(* IEC 61131-3 sources: vscode-structured-text/test/format/fixtures, 10 files *)

(* ---- types.expected.st ---- *)
TYPE tComplex
(*
Copyright ©<Company>. All rights reserved.
*)
    STRUCT
        rRe : Real; //Complex real part
        rIm : Real; //Complex imaginary part
    END_STRUCT
END_TYPE

TYPE uMaCommand :
    UNION
        b : tMaCommand; //For Bit Access
        w : Word;       //For Word Access
    END_UNION
END_TYPE

TYPE eColor : (Red := 0, Green, Blue);
END_TYPE
TYPE tArr : Array[1..10] Of Pointer To Int;
END_TYPE

(* ---- types.input.st ---- *)
TYPE tComplex
(*
Copyright ©<Company>. All rights reserved.
*)
STRUCT
rRe : REAL ; //Complex real part
rIm : REAL ; //Complex imaginary part
END_STRUCT
END_TYPE

TYPE uMaCommand :
UNION
 b   : tMaCommand; //For Bit Access
 w   : WORD;  //For Word Access
END_UNION
END_TYPE

TYPE eColor : (Red := 0, Green, Blue); END_TYPE
TYPE tArr : ARRAY [1..10] OF POINTER TO INT; END_TYPE

(* ---- oneline.expected.st ---- *)
FUNCTION fcAdd : Int
VAR_INPUT
    a : Int;
    b : Int;
END_VAR
tiSourcIndex                            := tiSourcIndex + 1;
tiDestinationIndex                      := tiDestinationIndex + 1;
If xxx Then
    yyy                                 := 1;
End_If
fcAdd                                   := a + b;
END_FUNCTION

(* ---- oneline.input.st ---- *)
FUNCTION fcAdd : INT
VAR_INPUT a : INT; b : INT; END_VAR
tiSourcIndex := tiSourcIndex + 1; tiDestinationIndex := tiDestinationIndex + 1;
IF xxx THEN yyy := 1; END_IF
fcAdd:=a+b;
END_FUNCTION

(* ---- fbruntime.expected.st ---- *)
(*

**©2026 <Company> - TITLE =[V#01.01.01.03] Measures task runtime and jitter**

========================  ================  ===========  =========================================
Version Number            Date              Signature    Description
========================  ================  ===========  =========================================
V#01.01.01.03             2026.06.01        <Sign>         Original version.
========================  ================  ===========  =========================================
*)

FUNCTION_BLOCK fbRuntime
(*
Copyright ©2026 <Company>. All rights reserved.
AUTHOR : <Sign>
FAMILY : System
NAME   : fbRuntime
*)

VAR CONSTANT
    {attribute 'hide'} cliNsPerUs : LInt := 1000;      //Nanoseconds per microsecond
END_VAR

VAR_INPUT
    ibStart : Bool; //Start call
    ibReset : Bool; //Reset min and max
END_VAR

VAR_OUTPUT
    qltRuntime       : LTime; // Actual runtime
    qliRuntimeJitter : LInt;  // [us] Runtime jitter
    qltRuntimeMax    : LTime; // Maximum runtime
    qltRuntimemin    : LTime; // Minimum runtime
END_VAR

VAR //Static
    {attribute 'hide'} sltNow        : LTime;
    {attribute 'hide'} sltRuntimeMax : LTime;
END_VAR

VAR_TEMP
    {attribute 'hide'} tbRestart  : Bool;
    {attribute 'hide'} tltRuntime : LTime;
    {attribute 'hide'} tliJitter  : LInt;
    {attribute 'hide'} tltNow     : LTime;
END_VAR

//Populate Temporaries
tbRestart                               := gSystem.bRestart();
tltNow                                  := LTime();
tltRuntime                              := tltNow - sltNow;

//Handle restart and reset
If (ibReset Or tbRestart) Then
    sltRuntimeMax                       := LTime#0s;
    sltRuntimeMin                       := LTime#1d;
    sltNow                              := tltNow;
    Return;
End_If;

//Handle start and end call
If ibStart Then
    sltNow                              := tltNow;
    qltRuntime                          := Ltime#0s;
    qliRuntimeJitter                    := 0;
    Return;
End_If;

//Handle Min/Max cycle time
If (tltRuntime > sltRuntimeMax) Then
    sltRuntimeMax                       := tltRuntime;
Elsif (tltRuntime < sltRuntimeMin) Then
    sltRuntimeMin                       := tltRuntime;
End_If;
tliJitter                               := (LTime_To_LInt(tltRuntime) - sliJitter) / cliNsPerUs;
sliJitter                               := LTime_To_LInt(tltRuntime);

//Write to outputs
qltRuntime                              := tltRuntime;
qliRuntimeJitter                        := tliJitter; // jitter
qltRuntimeMax                           := sltRuntimeMax;
qltRuntimeMin                           := sltRuntimeMin;
END_FUNCTION_BLOCK

(* ---- fbruntime.input.st ---- *)
(*

**©2026 <Company> - TITLE =[V#01.01.01.03] Measures task runtime and jitter**

========================  ================  ===========  =========================================
Version Number            Date              Signature    Description
========================  ================  ===========  =========================================
V#01.01.01.03             2026.06.01        <Sign>         Original version.
========================  ================  ===========  =========================================
*)

FUNCTION_BLOCK fbRuntime
(*
Copyright ©2026 <Company>. All rights reserved.
AUTHOR : <Sign>
FAMILY : System
NAME   : fbRuntime
*)

VAR CONSTANT
{attribute 'hide'}     cliNsPerUs : Lint:= 1000;      //Nanoseconds per microsecond
END_VAR
VAR_INPUT
 ibStart    : Bool;        //Start call
 ibReset    : Bool;        //Reset min and max
END_VAR

VAR_OUTPUT
 qltRuntime   : LTime;  // Actual runtime
 qliRuntimeJitter  : Lint;         // [us] Runtime jitter
 qltRuntimeMax   : LTime;  // Maximum runtime
 qltRuntimemin   : LTime;  // Minimum runtime
END_VAR

VAR //Static
{attribute 'hide'}     sltNow  : LTime;
{attribute 'hide'}     sltRuntimeMax : LTime;
END_VAR

VAR_TEMP
{attribute 'hide'}     tbRestart : Bool;
{attribute 'hide'}     tltRuntime    : LTime;
{attribute 'hide'}     tliJitter    : Lint ;
{attribute 'hide'}     tltNow  : LTime;
END_VAR

//Populate Temporaries
tbRestart := gSystem.bRestart();
tltNow  := LTime();
tltRuntime := tltNow - sltNow;

//Handle restart and reset
IF (ibReset OR tbRestart) THEN
sltRuntimeMax := LTime#0s;
    sltRuntimeMin                  := LTime#1d;
      sltNow                        := tltNow;
    RETURN;
END_IF;

//Handle start and end call
If ibStart Then sltNow := tltNow; qltRuntime := Ltime#0s;
    qliRuntimeJitter            := 0;
    Return;
End_If;

//Handle Min/Max cycle time
If (tltRuntime > sltRuntimeMax) Then
    sltRuntimeMax                    := tltRuntime;
Elsif (tltRuntime < sltRuntimeMin) Then
    sltRuntimeMin                    := tltRuntime;
End_If;
tliJitter:=(LTIME_TO_LINT(tltRuntime)-sliJitter)/cliNsPerUs;
sliJitter                            := LTime_To_Lint(tltRuntime);

//Write to outputs
qltRuntime                          := tltRuntime;
qliRuntimeJitter            := tliJitter; // jitter
qltRuntimeMax              := sltRuntimeMax;
qltRuntimeMin               := sltRuntimeMin;
END_FUNCTION_BLOCK

(* ---- oop.expected.st ---- *)
{attribute 'qualified_only'}
INTERFACE iMotor EXTENDS iBase
METHOD mStart : Bool
VAR_INPUT
    ibForce : Bool;
END_VAR
END_METHOD
END_INTERFACE

FUNCTION_BLOCK PUBLIC fbMotor EXTENDS fbBase IMPLEMENTS iMotor
VAR_INPUT
    RX : Bool;   //Initialize filter
END_VAR;

VAR //Static Data
    sbRx   : Bool;   //Initialize filter
    sRef   : Reference To Int;
    spData : Pointer To tData;
END_VAR;

VAR_TEMP
    tbRx : Bool;    //Initialize filter
END_VAR;
BEGIN
tbRx                                    := RX And Not sbRx; //tbRx is positive edge for RX
sbRx                                    := RX;              //Save RX in sbRx to disable edge as long as RX stays true.
{IF defined (DEBUG)}
If tbRx Then
    This^.mLog(sMsg := 'edge');
End_If;
{END_IF}
spData                                  := __New(tData);
sRef REF= siValue;
If ((tbyXa And 16#01) <> 16#00) Then  //Test for positive edge on bit zero in the byte
    sbAlarm S= True;
End_If
METHOD PRIVATE mLog : Bool
VAR_INPUT
    sMsg : String(80);
END_VAR
mLog                                    := True;
END_METHOD

PROPERTY pbRunning : Bool
END_PROPERTY
END_FUNCTION_BLOCK

(* ---- oop.input.st ---- *)
{attribute 'qualified_only'}
INTERFACE iMotor EXTENDS iBase
METHOD mStart : BOOL
VAR_INPUT
ibForce : BOOL;
END_VAR
END_METHOD
END_INTERFACE

FUNCTION_BLOCK PUBLIC fbMotor EXTENDS fbBase IMPLEMENTS iMotor
VAR_INPUT
    RX   : Bool ;   //Initialize filter
END_VAR;
VAR //Static Data
    sbRx  : Bool ;   //Initialize filter
    sRef : REFERENCE TO INT;
    spData : POINTER TO tData;
END_VAR;
VAR_TEMP
    tbRx         : Bool ;    //Initialize filter
END_VAR;
BEGIN
tbRx   := RX And Not sbRx; //tbRx is positive edge for RX
sbRx   := RX;              //Save RX in sbRx to disable edge as long as RX stays true.
{IF defined (DEBUG)}
If tbRx Then
    THIS^.mLog(sMsg := 'edge');
End_If;
{END_IF}
spData := __NEW(tData);
sRef REF= siValue;
IF ((tbyXa AND 16#01) <> 16#00) THEN  //Test for positive edge on bit zero in the byte
    sbAlarm S= TRUE;
END_IF
METHOD PRIVATE mLog : BOOL
VAR_INPUT
    sMsg : STRING(80);
END_VAR
mLog := TRUE;
END_METHOD

PROPERTY pbRunning : BOOL
END_PROPERTY
END_FUNCTION_BLOCK

(* ---- fsm.expected.st ---- *)
VAR CONSTANT
    //State Machine Constants
    ciInitState   : Int := 00; //Initial State of Control Element
    ciLow         : Int := 01; //Control Element in Low state
    ciTransitHigh : Int := 02; //Control Element in transit to High state
END_VAR

VAR //Static
    siState : Int; //State of Equipment Under Control
END_VAR
//State machine
Case siState Of
    ciInitState: //Initial State of EUC
        If bHigh Then
            siState                     := ciHigh;
        Elsif bLow Then
            siState                     := ciLow;
        End_If
    // EUC in Low state
    ciLow:
        If bSwitch Then
            siState                     := ciTransitHigh;
        End_If
    ciTransitHigh, ciTransitLow:
        x                               := 1;
        y                               := 22;
    Else
        siState                         := ciInitState;
End_Case;
Repeat
    i                                   := i + 1;
Until i > 10
End_Repeat;
While a And
        b Do
    x                                   := -1;
End_While
For tiII := tiBufferLength - 1 To 1 By -1 Do
    srBuffer[tiII + 1]                  := srBuffer[tiII];
End_For;

(* ---- fsm.input.st ---- *)
VAR CONSTANT
//State Machine Constants
ciInitState : INT := 00; //Initial State of Control Element
ciLow : INT := 01; //Control Element in Low state
ciTransitHigh : INT := 02; //Control Element in transit to High state
END_VAR
VAR //Static
siState : INT ; //State of Equipment Under Control
END_VAR
//State machine
CASE siState OF
ciInitState : //Initial State of EUC
IF bHigh THEN siState := ciHigh; ELSIF bLow THEN siState := ciLow; END_IF
// EUC in Low state
ciLow: IF bSwitch THEN
siState:=ciTransitHigh;
END_IF
ciTransitHigh, ciTransitLow:
x := 1; y := 22;
ELSE
siState := ciInitState;
END_CASE;
REPEAT i := i + 1; UNTIL i > 10 END_REPEAT;
WHILE a AND
    b DO x := -1; END_WHILE
FOR tiII := tiBufferLength - 1 TO 1 BY -1 DO srBuffer[tiII + 1] := srBuffer[tiII]; END_FOR;
